(* IEC 61131-3 sources: NachHouse_TST/ROOM_API_PILOT/CODEX_BACKUP_BEFORE_SK_COMMENTS_20260826_2356, 11 files *)

(* ---- 02_TYPES.ST ---- *)
(* ROOM_API_PILOT - logical API and transport types. *)

TYPE T_API_COMMAND_RESULT :
STRUCT
    ClientId       : STRING[36];
    RequestId      : UDINT;
    Result         : USINT;
    Message        : STRING[80];
    ConfigRevision : UDINT;
    StateRevision  : UDINT;
END_STRUCT
END_TYPE

TYPE T_API_INFO :
STRUCT
    ApiVersion        : STRING[32];
    ConfigRevision    : UDINT;
    StateRevision     : UDINT;
    MaxRooms          : USINT;
    LastCommandResult : T_API_COMMAND_RESULT;
END_STRUCT
END_TYPE

TYPE T_ROOM_CONFIG :
STRUCT
    Used        : BOOL;
    RoomId      : UDINT;
    Name        : STRING[64];
    ProjectName : STRING[64];
    IconId      : UINT;
    SortDefault : UINT;
END_STRUCT
END_TYPE

TYPE T_API_CONFIG :
STRUCT
    Rooms : ARRAY[1..40] OF T_ROOM_CONFIG;
END_STRUCT
END_TYPE

TYPE T_ROOM_STATE :
STRUCT
    RoomId       : UDINT;
    Temperature  : REAL;
    Humidity     : REAL;
    Presence     : BOOL;
    DayPhase     : UINT;
    CategoryMask : DWORD;
    AlarmLevel   : USINT;
    Online       : BOOL;
END_STRUCT
END_TYPE

TYPE T_API_STATE :
STRUCT
    Rooms : ARRAY[1..40] OF T_ROOM_STATE;
END_STRUCT
END_TYPE

TYPE T_API_COMMAND_ROOM :
STRUCT
    ClientId     : STRING[36];
    RequestId    : UDINT;
    Action       : USINT;
    RoomId       : UDINT;
    SourceRoomId : UDINT;
    Name         : STRING[64];
    ProjectName  : STRING[64];
END_STRUCT
END_TYPE

TYPE T_API_CONFIG_CHANGE :
STRUCT
    Valid     : BOOL;
    Operation : USINT;
    RoomId    : UDINT;
    Room      : T_ROOM_CONFIG;
END_STRUCT
END_TYPE

TYPE T_API_STATE_CHANGE :
STRUCT
    Valid     : BOOL;
    Operation : USINT;
    RoomId    : UDINT;
    Room      : T_ROOM_STATE;
END_STRUCT
END_TYPE

TYPE T_API_CONFIG_DIFF :
STRUCT
    Valid        : BOOL;
    FromRevision : UDINT;
    ToRevision   : UDINT;
    FullRequired : BOOL;
    ChangeCount  : USINT;
    Changes      : ARRAY[1..40] OF T_API_CONFIG_CHANGE;
END_STRUCT
END_TYPE

TYPE T_API_STATE_DIFF :
STRUCT
    Valid        : BOOL;
    FromRevision : UDINT;
    ToRevision   : UDINT;
    FullRequired : BOOL;
    ChangeCount  : USINT;
    Changes      : ARRAY[1..40] OF T_API_STATE_CHANGE;
END_STRUCT
END_TYPE

(* Transport handshake used to retrieve one retained diff frame. *)
TYPE T_API_SYNC_REQUEST :
STRUCT
    ClientId           : STRING[36];
    RequestId          : UDINT;
    ConfigFromRevision : UDINT;
    StateFromRevision  : UDINT;
END_STRUCT
END_TYPE

TYPE T_API_SYNC_RESPONSE :
STRUCT
    ClientId   : STRING[36];
    RequestId  : UDINT;
    Result     : USINT;
    Message    : STRING[80];
    ConfigMode : USINT;
    StateMode  : USINT;
    ConfigDiff : T_API_CONFIG_DIFF;
    StateDiff  : T_API_STATE_DIFF;
END_STRUCT
END_TYPE

(* Manual test input. It is deliberately separate from ApiCommand.Room. *)
TYPE T_API_TEST_STATE_REQUEST :
STRUCT
    ClientId     : STRING[36];
    RequestId    : UDINT;
    RoomId       : UDINT;
    Temperature  : REAL;
    Humidity     : REAL;
    Presence     : BOOL;
    DayPhase     : UINT;
    CategoryMask : DWORD;
    AlarmLevel   : USINT;
    Online       : BOOL;
END_STRUCT
END_TYPE

(* ---- 01_CONSTANTS.ST ---- *)
(* ROOM_API_PILOT - public numeric contract and limits. *)

VAR_GLOBAL CONSTANT
    C_API_VERSION          : STRING[32] := 'ROOM_API_PILOT/1';
    C_MAX_ROOMS            : USINT := 40;
    C_DIFF_HISTORY_DEPTH   : USINT := 8;

    API_ACTION_NONE          : USINT := 0;
    API_ACTION_ADD_ROOM      : USINT := 1;
    API_ACTION_DELETE_ROOM   : USINT := 2;
    API_ACTION_COPY_ROOM     : USINT := 3;
    API_ACTION_SET_ROOM_DATA : USINT := 4;

    API_RESULT_NONE               : USINT := 0;
    API_RESULT_OK                 : USINT := 1;
    API_RESULT_ERROR              : USINT := 2;
    API_RESULT_NOT_FOUND          : USINT := 3;
    API_RESULT_NO_FREE_SLOT       : USINT := 4;
    API_RESULT_ALREADY_EXISTS     : USINT := 5;
    API_RESULT_INVALID_ARGUMENT   : USINT := 6;
    API_RESULT_UNSUPPORTED_ACTION : USINT := 7;

    API_DIFF_NONE   : USINT := 0;
    API_DIFF_UPSERT : USINT := 1;
    API_DIFF_DELETE : USINT := 2;

    API_SYNC_CURRENT       : USINT := 0;
    API_SYNC_DIFF          : USINT := 1;
    API_SYNC_FULL_REQUIRED : USINT := 2;

    API_ALARM_OK      : USINT := 0;
    API_ALARM_WARNING : USINT := 1;
    API_ALARM_ALARM   : USINT := 2;

    API_DAY_PHASE_DAY   : UINT := 140;
    API_DAY_PHASE_DUSK  : UINT := 142;
    API_DAY_PHASE_NIGHT : UINT := 144;
    API_DAY_PHASE_DAWN  : UINT := 146;

    API_DEFAULT_ICON_ID     : UINT := 16;
    API_DEFAULT_TEMPERATURE : REAL := 20.0;
    API_DEFAULT_HUMIDITY    : REAL := 40.0;
END_VAR

(* ---- 03_PUBLIC_API.ST ---- *)
(*
   All client-visible objects are global and marked PUBLIC_API.
   The client must write request payload fields first and Execute last.
   Snapshot objects ApiConfig and ApiState are read-only by contract.
*)

VAR_GLOBAL
    ApiInfo       {PUBLIC_API} : T_API_INFO;
    ApiConfig     {PUBLIC_API} : T_API_CONFIG;
    ApiState      {PUBLIC_API} : T_API_STATE;

    ApiConfigDiff {PUBLIC_API} : T_API_CONFIG_DIFF;
    ApiStateDiff  {PUBLIC_API} : T_API_STATE_DIFF;

    ApiCommandRoom     {PUBLIC_API} : T_API_COMMAND_ROOM;
    ApiCommandExecute  {PUBLIC_API} : BOOL;
    ApiCommandBusy     {PUBLIC_API} : BOOL;
    ApiCommandFinished {PUBLIC_API} : BOOL;
    ApiCommandResult   {PUBLIC_API} : T_API_COMMAND_RESULT;

    ApiSyncRequest  {PUBLIC_API} : T_API_SYNC_REQUEST;
    ApiSyncExecute  {PUBLIC_API} : BOOL;
    ApiSyncBusy     {PUBLIC_API} : BOOL;
    ApiSyncFinished {PUBLIC_API} : BOOL;
    ApiSyncResponse {PUBLIC_API} : T_API_SYNC_RESPONSE;

    ApiTestStateRequest  {PUBLIC_API} : T_API_TEST_STATE_REQUEST;
    ApiTestStateExecute  {PUBLIC_API} : BOOL;
    ApiTestStateBusy     {PUBLIC_API} : BOOL;
    ApiTestStateFinished {PUBLIC_API} : BOOL;
    ApiTestStateResult   {PUBLIC_API} : T_API_COMMAND_RESULT;
END_VAR

(* ---- 04_INTERNAL.ST ---- *)
(* Internal state is not exported to TecoApi / PLCComS. *)

VAR_GLOBAL
    ApiInitialized : BOOL;

    ApiConfigShadow : ARRAY[1..40] OF T_ROOM_CONFIG;
    ApiStateShadow  : ARRAY[1..40] OF T_ROOM_STATE;

    ApiConfigDiffHistory : ARRAY[1..8] OF T_API_CONFIG_DIFF;
    ApiStateDiffHistory  : ARRAY[1..8] OF T_API_STATE_DIFF;
    ApiConfigHistoryHead : USINT;
    ApiStateHistoryHead  : USINT;

    ApiLastCommandClientId  : STRING[36];
    ApiLastCommandRequestId : UDINT;
    ApiLastStoredResult     : T_API_COMMAND_RESULT;
END_VAR

(* ---- 05_UTILS.ST ---- *)
(* ROOM_API_PILOT - small deterministic helpers. *)

FUNCTION ApiRoomConfigEqual : BOOL
VAR_INPUT
    A : T_ROOM_CONFIG;
    B : T_ROOM_CONFIG;
END_VAR

ApiRoomConfigEqual :=
    (A.Used = B.Used) AND
    (A.RoomId = B.RoomId) AND
    (A.Name = B.Name) AND
    (A.ProjectName = B.ProjectName) AND
    (A.IconId = B.IconId) AND
    (A.SortDefault = B.SortDefault);
END_FUNCTION

FUNCTION ApiRoomStateEqual : BOOL
VAR_INPUT
    A : T_ROOM_STATE;
    B : T_ROOM_STATE;
END_VAR

ApiRoomStateEqual :=
    (A.RoomId = B.RoomId) AND
    (A.Temperature = B.Temperature) AND
    (A.Humidity = B.Humidity) AND
    (A.Presence = B.Presence) AND
    (A.DayPhase = B.DayPhase) AND
    (A.CategoryMask = B.CategoryMask) AND
    (A.AlarmLevel = B.AlarmLevel) AND
    (A.Online = B.Online);
END_FUNCTION

FUNCTION ApiFindConfigSlot : USINT
VAR_INPUT
    RoomId : UDINT;
END_VAR
VAR
    i : USINT;
END_VAR

ApiFindConfigSlot := 0;
IF RoomId <> 0 THEN
    FOR i := 1 TO C_MAX_ROOMS DO
        IF ApiConfig.Rooms[i].Used AND (ApiConfig.Rooms[i].RoomId = RoomId) THEN
            ApiFindConfigSlot := i;
            RETURN;
        END_IF;
    END_FOR;
END_IF;
END_FUNCTION

FUNCTION ApiFindStateSlot : USINT
VAR_INPUT
    RoomId : UDINT;
END_VAR
VAR
    i : USINT;
END_VAR

ApiFindStateSlot := 0;
IF RoomId <> 0 THEN
    FOR i := 1 TO C_MAX_ROOMS DO
        IF ApiState.Rooms[i].RoomId = RoomId THEN
            ApiFindStateSlot := i;
            RETURN;
        END_IF;
    END_FOR;
END_IF;
END_FUNCTION

FUNCTION ApiFindFreeConfigSlot : USINT
VAR
    i : USINT;
END_VAR

ApiFindFreeConfigSlot := 0;
FOR i := 1 TO C_MAX_ROOMS DO
    IF NOT ApiConfig.Rooms[i].Used THEN
        ApiFindFreeConfigSlot := i;
        RETURN;
    END_IF;
END_FOR;
END_FUNCTION

FUNCTION ApiFindFreeStateSlot : USINT
VAR
    i : USINT;
END_VAR

ApiFindFreeStateSlot := 0;
FOR i := 1 TO C_MAX_ROOMS DO
    IF ApiState.Rooms[i].RoomId = 0 THEN
        ApiFindFreeStateSlot := i;
        RETURN;
    END_IF;
END_FOR;
END_FUNCTION

FUNCTION ApiClearRoomConfig : BOOL
VAR_IN_OUT
    Room : T_ROOM_CONFIG;
END_VAR

Room.Used := FALSE;
Room.RoomId := 0;
Room.Name := '';
Room.ProjectName := '';
Room.IconId := 0;
Room.SortDefault := 0;
ApiClearRoomConfig := TRUE;
END_FUNCTION

FUNCTION ApiClearRoomState : BOOL
VAR_IN_OUT
    Room : T_ROOM_STATE;
END_VAR

Room.RoomId := 0;
Room.Temperature := 0.0;
Room.Humidity := 0.0;
Room.Presence := FALSE;
Room.DayPhase := API_DAY_PHASE_DAY;
Room.CategoryMask := DWORD#16#00000000;
Room.AlarmLevel := API_ALARM_OK;
Room.Online := FALSE;
ApiClearRoomState := TRUE;
END_FUNCTION

FUNCTION ApiClearConfigDiff : BOOL
VAR_IN_OUT
    Diff : T_API_CONFIG_DIFF;
END_VAR
VAR
    i : USINT;
END_VAR

Diff.Valid := FALSE;
Diff.FromRevision := 0;
Diff.ToRevision := 0;
Diff.FullRequired := FALSE;
Diff.ChangeCount := 0;
FOR i := 1 TO C_MAX_ROOMS DO
    Diff.Changes[i].Valid := FALSE;
    Diff.Changes[i].Operation := API_DIFF_NONE;
    Diff.Changes[i].RoomId := 0;
    ApiClearRoomConfig(Diff.Changes[i].Room);
END_FOR;
ApiClearConfigDiff := TRUE;
END_FUNCTION

FUNCTION ApiClearStateDiff : BOOL
VAR_IN_OUT
    Diff : T_API_STATE_DIFF;
END_VAR
VAR
    i : USINT;
END_VAR

Diff.Valid := FALSE;
Diff.FromRevision := 0;
Diff.ToRevision := 0;
Diff.FullRequired := FALSE;
Diff.ChangeCount := 0;
FOR i := 1 TO C_MAX_ROOMS DO
    Diff.Changes[i].Valid := FALSE;
    Diff.Changes[i].Operation := API_DIFF_NONE;
    Diff.Changes[i].RoomId := 0;
    ApiClearRoomState(Diff.Changes[i].Room);
END_FOR;
ApiClearStateDiff := TRUE;
END_FUNCTION

FUNCTION ApiNextRevision : UDINT
VAR_INPUT
    Revision : UDINT;
END_VAR

ApiNextRevision := Revision + 1;
IF ApiNextRevision = 0 THEN
    ApiNextRevision := 1;
END_IF;
END_FUNCTION

FUNCTION ApiValidDayPhase : BOOL
VAR_INPUT
    DayPhase : UINT;
END_VAR

ApiValidDayPhase :=
    (DayPhase = API_DAY_PHASE_DAY) OR
    (DayPhase = API_DAY_PHASE_DUSK) OR
    (DayPhase = API_DAY_PHASE_NIGHT) OR
    (DayPhase = API_DAY_PHASE_DAWN);
END_FUNCTION

(* ---- 06_DIFF_ENGINE.ST ---- *)
(*
   Diff engine.
   One PLC transaction creates one revision and one complete diff frame.
   Eight frames are retained. A client asks for one next frame at a time.
*)

FUNCTION ApiCaptureConfigChanges : BOOL
VAR
    i          : USINT;
    count      : USINT;
    oldRev     : UDINT;
    newRev     : UDINT;
    anyChanged : BOOL;
END_VAR

anyChanged := FALSE;
FOR i := 1 TO C_MAX_ROOMS DO
    IF NOT ApiRoomConfigEqual(ApiConfig.Rooms[i], ApiConfigShadow[i]) THEN
        anyChanged := TRUE;
    END_IF;
END_FOR;

ApiCaptureConfigChanges := anyChanged;
IF NOT anyChanged THEN
    RETURN;
END_IF;

ApiClearConfigDiff(ApiConfigDiff);
oldRev := ApiInfo.ConfigRevision;
newRev := ApiNextRevision(oldRev);
ApiConfigDiff.FromRevision := oldRev;
ApiConfigDiff.ToRevision := newRev;
ApiConfigDiff.FullRequired := FALSE;
count := 0;

FOR i := 1 TO C_MAX_ROOMS DO
    IF NOT ApiRoomConfigEqual(ApiConfig.Rooms[i], ApiConfigShadow[i]) THEN
        count := count + 1;
        ApiConfigDiff.Changes[count].Valid := TRUE;

        IF ApiConfig.Rooms[i].Used THEN
            ApiConfigDiff.Changes[count].Operation := API_DIFF_UPSERT;
            ApiConfigDiff.Changes[count].RoomId := ApiConfig.Rooms[i].RoomId;
            ApiConfigDiff.Changes[count].Room := ApiConfig.Rooms[i];
        ELSE
            ApiConfigDiff.Changes[count].Operation := API_DIFF_DELETE;
            ApiConfigDiff.Changes[count].RoomId := ApiConfigShadow[i].RoomId;
            ApiClearRoomConfig(ApiConfigDiff.Changes[count].Room);
        END_IF;
    END_IF;

    ApiConfigShadow[i] := ApiConfig.Rooms[i];
END_FOR;

ApiConfigDiff.ChangeCount := count;
ApiConfigDiff.Valid := TRUE;
ApiInfo.ConfigRevision := newRev;

IF ApiConfigHistoryHead >= C_DIFF_HISTORY_DEPTH THEN
    ApiConfigHistoryHead := 1;
ELSE
    ApiConfigHistoryHead := ApiConfigHistoryHead + 1;
END_IF;
ApiConfigDiffHistory[ApiConfigHistoryHead] := ApiConfigDiff;
END_FUNCTION

FUNCTION ApiCaptureStateChanges : BOOL
VAR
    i          : USINT;
    count      : USINT;
    oldRev     : UDINT;
    newRev     : UDINT;
    anyChanged : BOOL;
END_VAR

anyChanged := FALSE;
FOR i := 1 TO C_MAX_ROOMS DO
    IF NOT ApiRoomStateEqual(ApiState.Rooms[i], ApiStateShadow[i]) THEN
        anyChanged := TRUE;
    END_IF;
END_FOR;

ApiCaptureStateChanges := anyChanged;
IF NOT anyChanged THEN
    RETURN;
END_IF;

ApiClearStateDiff(ApiStateDiff);
oldRev := ApiInfo.StateRevision;
newRev := ApiNextRevision(oldRev);
ApiStateDiff.FromRevision := oldRev;
ApiStateDiff.ToRevision := newRev;
ApiStateDiff.FullRequired := FALSE;
count := 0;

FOR i := 1 TO C_MAX_ROOMS DO
    IF NOT ApiRoomStateEqual(ApiState.Rooms[i], ApiStateShadow[i]) THEN
        count := count + 1;
        ApiStateDiff.Changes[count].Valid := TRUE;

        IF ApiState.Rooms[i].RoomId <> 0 THEN
            ApiStateDiff.Changes[count].Operation := API_DIFF_UPSERT;
            ApiStateDiff.Changes[count].RoomId := ApiState.Rooms[i].RoomId;
            ApiStateDiff.Changes[count].Room := ApiState.Rooms[i];
        ELSE
            ApiStateDiff.Changes[count].Operation := API_DIFF_DELETE;
            ApiStateDiff.Changes[count].RoomId := ApiStateShadow[i].RoomId;
            ApiClearRoomState(ApiStateDiff.Changes[count].Room);
        END_IF;
    END_IF;

    ApiStateShadow[i] := ApiState.Rooms[i];
END_FOR;

ApiStateDiff.ChangeCount := count;
ApiStateDiff.Valid := TRUE;
ApiInfo.StateRevision := newRev;

IF ApiStateHistoryHead >= C_DIFF_HISTORY_DEPTH THEN
    ApiStateHistoryHead := 1;
ELSE
    ApiStateHistoryHead := ApiStateHistoryHead + 1;
END_IF;
ApiStateDiffHistory[ApiStateHistoryHead] := ApiStateDiff;
END_FUNCTION

(* ---- 07_INIT.ST ---- *)
(* Cold-start initialization and deterministic pilot data. *)

FUNCTION ApiPilotInit : BOOL
VAR
    i : USINT;
END_VAR

ApiPilotInit := ApiInitialized;
IF ApiInitialized THEN
    RETURN;
END_IF;

FOR i := 1 TO C_MAX_ROOMS DO
    ApiClearRoomConfig(ApiConfig.Rooms[i]);
    ApiClearRoomState(ApiState.Rooms[i]);
    ApiClearRoomConfig(ApiConfigShadow[i]);
    ApiClearRoomState(ApiStateShadow[i]);
END_FOR;

FOR i := 1 TO C_DIFF_HISTORY_DEPTH DO
    ApiClearConfigDiff(ApiConfigDiffHistory[i]);
    ApiClearStateDiff(ApiStateDiffHistory[i]);
END_FOR;

(* Four sample rooms. Values are test data only. *)
ApiConfig.Rooms[1].Used := TRUE;
ApiConfig.Rooms[1].RoomId := 1;
ApiConfig.Rooms[1].Name := 'Obyvacka';
ApiConfig.Rooms[1].ProjectName := '1.01';
ApiConfig.Rooms[1].IconId := 16;
ApiConfig.Rooms[1].SortDefault := 1;

ApiConfig.Rooms[2].Used := TRUE;
ApiConfig.Rooms[2].RoomId := 2;
ApiConfig.Rooms[2].Name := 'Kuchyna';
ApiConfig.Rooms[2].ProjectName := '1.07';
ApiConfig.Rooms[2].IconId := 16;
ApiConfig.Rooms[2].SortDefault := 2;

ApiConfig.Rooms[3].Used := TRUE;
ApiConfig.Rooms[3].RoomId := 3;
ApiConfig.Rooms[3].Name := 'Spalna';
ApiConfig.Rooms[3].ProjectName := '1.09';
ApiConfig.Rooms[3].IconId := 16;
ApiConfig.Rooms[3].SortDefault := 3;

ApiConfig.Rooms[4].Used := TRUE;
ApiConfig.Rooms[4].RoomId := 4;
ApiConfig.Rooms[4].Name := 'Terasa';
ApiConfig.Rooms[4].ProjectName := 'E.01';
ApiConfig.Rooms[4].IconId := 19;
ApiConfig.Rooms[4].SortDefault := 4;

ApiState.Rooms[1].RoomId := 1;
ApiState.Rooms[1].Temperature := 22.5;
ApiState.Rooms[1].Humidity := 45.0;
ApiState.Rooms[1].Presence := TRUE;
ApiState.Rooms[1].DayPhase := API_DAY_PHASE_DAY;
ApiState.Rooms[1].CategoryMask := DWORD#16#00000007;
ApiState.Rooms[1].AlarmLevel := API_ALARM_OK;
ApiState.Rooms[1].Online := TRUE;

ApiState.Rooms[2].RoomId := 2;
ApiState.Rooms[2].Temperature := 23.0;
ApiState.Rooms[2].Humidity := 48.0;
ApiState.Rooms[2].Presence := FALSE;
ApiState.Rooms[2].DayPhase := API_DAY_PHASE_DUSK;
ApiState.Rooms[2].CategoryMask := DWORD#16#00000003;
ApiState.Rooms[2].AlarmLevel := API_ALARM_WARNING;
ApiState.Rooms[2].Online := TRUE;

ApiState.Rooms[3].RoomId := 3;
ApiState.Rooms[3].Temperature := 21.8;
ApiState.Rooms[3].Humidity := 42.0;
ApiState.Rooms[3].Presence := TRUE;
ApiState.Rooms[3].DayPhase := API_DAY_PHASE_NIGHT;
ApiState.Rooms[3].CategoryMask := DWORD#16#00000001;
ApiState.Rooms[3].AlarmLevel := API_ALARM_OK;
ApiState.Rooms[3].Online := TRUE;

ApiState.Rooms[4].RoomId := 4;
ApiState.Rooms[4].Temperature := 18.4;
ApiState.Rooms[4].Humidity := 58.0;
ApiState.Rooms[4].Presence := FALSE;
ApiState.Rooms[4].DayPhase := API_DAY_PHASE_DAWN;
ApiState.Rooms[4].CategoryMask := DWORD#16#00000004;
ApiState.Rooms[4].AlarmLevel := API_ALARM_ALARM;
ApiState.Rooms[4].Online := FALSE;

FOR i := 1 TO C_MAX_ROOMS DO
    ApiConfigShadow[i] := ApiConfig.Rooms[i];
    ApiStateShadow[i] := ApiState.Rooms[i];
END_FOR;

ApiInfo.ApiVersion := C_API_VERSION;
ApiInfo.ConfigRevision := 1;
ApiInfo.StateRevision := 1;
ApiInfo.MaxRooms := C_MAX_ROOMS;
ApiInfo.LastCommandResult.ClientId := '';
ApiInfo.LastCommandResult.RequestId := 0;
ApiInfo.LastCommandResult.Result := API_RESULT_NONE;
ApiInfo.LastCommandResult.Message := 'Ziadny prikaz';
ApiInfo.LastCommandResult.ConfigRevision := 1;
ApiInfo.LastCommandResult.StateRevision := 1;

ApiClearConfigDiff(ApiConfigDiff);
ApiConfigDiff.Valid := TRUE;
ApiConfigDiff.FromRevision := 0;
ApiConfigDiff.ToRevision := 1;
ApiConfigDiff.FullRequired := TRUE;

ApiClearStateDiff(ApiStateDiff);
ApiStateDiff.Valid := TRUE;
ApiStateDiff.FromRevision := 0;
ApiStateDiff.ToRevision := 1;
ApiStateDiff.FullRequired := TRUE;

ApiCommandRoom.ClientId := '';
ApiCommandRoom.RequestId := 0;
ApiCommandRoom.Action := API_ACTION_NONE;
ApiCommandRoom.RoomId := 0;
ApiCommandRoom.SourceRoomId := 0;
ApiCommandRoom.Name := '';
ApiCommandRoom.ProjectName := '';
ApiCommandExecute := FALSE;
ApiCommandBusy := FALSE;
ApiCommandFinished := FALSE;
ApiCommandResult := ApiInfo.LastCommandResult;

ApiSyncExecute := FALSE;
ApiSyncBusy := FALSE;
ApiSyncFinished := FALSE;
ApiTestStateExecute := FALSE;
ApiTestStateBusy := FALSE;
ApiTestStateFinished := FALSE;

ApiConfigHistoryHead := 0;
ApiStateHistoryHead := 0;
ApiLastCommandClientId := '';
ApiLastCommandRequestId := 0;
ApiLastStoredResult := ApiInfo.LastCommandResult;

ApiInitialized := TRUE;
ApiPilotInit := TRUE;
END_FUNCTION

(* ---- 08_COMMAND_ENGINE.ST ---- *)
(* ADD / DELETE / COPY / SET command processor. *)

FUNCTION ApiProcessRoomCommand : BOOL
VAR
    i             : USINT;
    configSlot    : USINT;
    stateSlot     : USINT;
    sourceCfgSlot : USINT;
    sourceStSlot  : USINT;
    maxSort       : UINT;
    sourceSort    : UINT;
    resultCode    : USINT;
    resultMessage : STRING[80];
    executeChange : BOOL;
END_VAR

ApiProcessRoomCommand := FALSE;
IF NOT ApiCommandExecute THEN
    RETURN;
END_IF;

ApiProcessRoomCommand := TRUE;
ApiCommandBusy := TRUE;
ApiCommandFinished := FALSE;

(* Exact retry of the latest command is idempotent. *)
IF (ApiCommandRoom.ClientId = ApiLastCommandClientId) AND
   (ApiCommandRoom.RequestId = ApiLastCommandRequestId) AND
   (ApiCommandRoom.RequestId <> 0) THEN

    ApiCommandResult := ApiLastStoredResult;
    ApiInfo.LastCommandResult := ApiLastStoredResult;

ELSE
    resultCode := API_RESULT_OK;
    resultMessage := 'OK';
    executeChange := FALSE;

    IF (ApiCommandRoom.ClientId = '') OR (ApiCommandRoom.RequestId = 0) THEN
        resultCode := API_RESULT_INVALID_ARGUMENT;
        resultMessage := 'Neplatny ClientId alebo RequestId';
    ELSE
        CASE ApiCommandRoom.Action OF

            API_ACTION_ADD_ROOM:
                IF (ApiCommandRoom.RoomId = 0) OR (ApiCommandRoom.Name = '') THEN
                    resultCode := API_RESULT_INVALID_ARGUMENT;
                    resultMessage := 'Neplatne ID alebo nazov';
                ELSIF ApiFindConfigSlot(ApiCommandRoom.RoomId) <> 0 THEN
                    resultCode := API_RESULT_ALREADY_EXISTS;
                    resultMessage := 'RoomId uz existuje';
                ELSE
                    configSlot := ApiFindFreeConfigSlot();
                    stateSlot := ApiFindFreeStateSlot();
                    IF (configSlot = 0) OR (stateSlot = 0) THEN
                        resultCode := API_RESULT_NO_FREE_SLOT;
                        resultMessage := 'Nie je volny slot';
                    ELSE
                        maxSort := 0;
                        FOR i := 1 TO C_MAX_ROOMS DO
                            IF ApiConfig.Rooms[i].Used AND
                               (ApiConfig.Rooms[i].SortDefault > maxSort) THEN
                                maxSort := ApiConfig.Rooms[i].SortDefault;
                            END_IF;
                        END_FOR;

                        ApiClearRoomConfig(ApiConfig.Rooms[configSlot]);
                        ApiConfig.Rooms[configSlot].Used := TRUE;
                        ApiConfig.Rooms[configSlot].RoomId := ApiCommandRoom.RoomId;
                        ApiConfig.Rooms[configSlot].Name := ApiCommandRoom.Name;
                        ApiConfig.Rooms[configSlot].ProjectName := ApiCommandRoom.ProjectName;
                        ApiConfig.Rooms[configSlot].IconId := API_DEFAULT_ICON_ID;
                        ApiConfig.Rooms[configSlot].SortDefault := maxSort + 1;

                        ApiClearRoomState(ApiState.Rooms[stateSlot]);
                        ApiState.Rooms[stateSlot].RoomId := ApiCommandRoom.RoomId;
                        ApiState.Rooms[stateSlot].Temperature := API_DEFAULT_TEMPERATURE;
                        ApiState.Rooms[stateSlot].Humidity := API_DEFAULT_HUMIDITY;
                        ApiState.Rooms[stateSlot].Presence := FALSE;
                        ApiState.Rooms[stateSlot].DayPhase := API_DAY_PHASE_DAY;
                        ApiState.Rooms[stateSlot].CategoryMask := DWORD#16#00000000;
                        ApiState.Rooms[stateSlot].AlarmLevel := API_ALARM_OK;
                        ApiState.Rooms[stateSlot].Online := TRUE;

                        executeChange := TRUE;
                        resultMessage := 'Miestnost pridana';
                    END_IF;
                END_IF;

            API_ACTION_DELETE_ROOM:
                configSlot := ApiFindConfigSlot(ApiCommandRoom.RoomId);
                stateSlot := ApiFindStateSlot(ApiCommandRoom.RoomId);
                IF (configSlot = 0) OR (stateSlot = 0) THEN
                    resultCode := API_RESULT_NOT_FOUND;
                    resultMessage := 'Miestnost nenajdena';
                ELSE
                    ApiClearRoomConfig(ApiConfig.Rooms[configSlot]);
                    ApiClearRoomState(ApiState.Rooms[stateSlot]);
                    executeChange := TRUE;
                    resultMessage := 'Miestnost zmazana';
                END_IF;

            API_ACTION_COPY_ROOM:
                sourceCfgSlot := ApiFindConfigSlot(ApiCommandRoom.SourceRoomId);
                sourceStSlot := ApiFindStateSlot(ApiCommandRoom.SourceRoomId);
                IF (ApiCommandRoom.RoomId = 0) OR
                   (ApiCommandRoom.RoomId = ApiCommandRoom.SourceRoomId) THEN
                    resultCode := API_RESULT_INVALID_ARGUMENT;
                    resultMessage := 'Neplatne cielove RoomId';
                ELSIF (sourceCfgSlot = 0) OR (sourceStSlot = 0) THEN
                    resultCode := API_RESULT_NOT_FOUND;
                    resultMessage := 'Zdrojova miestnost nenajdena';
                ELSIF ApiFindConfigSlot(ApiCommandRoom.RoomId) <> 0 THEN
                    resultCode := API_RESULT_ALREADY_EXISTS;
                    resultMessage := 'Cielove RoomId uz existuje';
                ELSE
                    configSlot := ApiFindFreeConfigSlot();
                    stateSlot := ApiFindFreeStateSlot();
                    IF (configSlot = 0) OR (stateSlot = 0) THEN
                        resultCode := API_RESULT_NO_FREE_SLOT;
                        resultMessage := 'Nie je volny slot';
                    ELSE
                        sourceSort := ApiConfig.Rooms[sourceCfgSlot].SortDefault;
                        FOR i := 1 TO C_MAX_ROOMS DO
                            IF ApiConfig.Rooms[i].Used AND
                               (ApiConfig.Rooms[i].SortDefault > sourceSort) THEN
                                ApiConfig.Rooms[i].SortDefault :=
                                    ApiConfig.Rooms[i].SortDefault + 1;
                            END_IF;
                        END_FOR;

                        ApiConfig.Rooms[configSlot] := ApiConfig.Rooms[sourceCfgSlot];
                        ApiConfig.Rooms[configSlot].RoomId := ApiCommandRoom.RoomId;
                        ApiConfig.Rooms[configSlot].SortDefault := sourceSort + 1;
                        IF ApiCommandRoom.Name <> '' THEN
                            ApiConfig.Rooms[configSlot].Name := ApiCommandRoom.Name;
                        END_IF;
                        IF ApiCommandRoom.ProjectName <> '' THEN
                            ApiConfig.Rooms[configSlot].ProjectName := ApiCommandRoom.ProjectName;
                        END_IF;

                        ApiState.Rooms[stateSlot] := ApiState.Rooms[sourceStSlot];
                        ApiState.Rooms[stateSlot].RoomId := ApiCommandRoom.RoomId;

                        executeChange := TRUE;
                        resultMessage := 'Miestnost skopirovana';
                    END_IF;
                END_IF;

            API_ACTION_SET_ROOM_DATA:
                configSlot := ApiFindConfigSlot(ApiCommandRoom.RoomId);
                IF configSlot = 0 THEN
                    resultCode := API_RESULT_NOT_FOUND;
                    resultMessage := 'Miestnost nenajdena';
                ELSIF ApiCommandRoom.Name = '' THEN
                    resultCode := API_RESULT_INVALID_ARGUMENT;
                    resultMessage := 'Nazov nesmie byt prazdny';
                ELSE
                    ApiConfig.Rooms[configSlot].Name := ApiCommandRoom.Name;
                    ApiConfig.Rooms[configSlot].ProjectName := ApiCommandRoom.ProjectName;
                    executeChange := TRUE;
                    resultMessage := 'Udaje miestnosti nastavene';
                END_IF;

            ELSE
                resultCode := API_RESULT_UNSUPPORTED_ACTION;
                resultMessage := 'Nepodporovana akcia';
        END_CASE;
    END_IF;

    IF executeChange AND (resultCode = API_RESULT_OK) THEN
        ApiCaptureConfigChanges();
        ApiCaptureStateChanges();
    END_IF;

    ApiCommandResult.ClientId := ApiCommandRoom.ClientId;
    ApiCommandResult.RequestId := ApiCommandRoom.RequestId;
    ApiCommandResult.Result := resultCode;
    ApiCommandResult.Message := resultMessage;
    ApiCommandResult.ConfigRevision := ApiInfo.ConfigRevision;
    ApiCommandResult.StateRevision := ApiInfo.StateRevision;

    ApiInfo.LastCommandResult := ApiCommandResult;
    ApiLastCommandClientId := ApiCommandRoom.ClientId;
    ApiLastCommandRequestId := ApiCommandRoom.RequestId;
    ApiLastStoredResult := ApiCommandResult;
END_IF;

ApiCommandExecute := FALSE;
ApiCommandBusy := FALSE;
ApiCommandFinished := TRUE;
END_FUNCTION

(* ---- 09_STATE_TEST.ST ---- *)
(* Manual, validated test-state writer. No real IO is connected. *)

FUNCTION ApiProcessTestState : BOOL
VAR
    configSlot    : USINT;
    stateSlot     : USINT;
    resultCode    : USINT;
    resultMessage : STRING[80];
END_VAR

ApiProcessTestState := FALSE;
IF NOT ApiTestStateExecute THEN
    RETURN;
END_IF;

ApiProcessTestState := TRUE;
ApiTestStateBusy := TRUE;
ApiTestStateFinished := FALSE;
resultCode := API_RESULT_OK;
resultMessage := 'Testovaci stav nastaveny';

configSlot := ApiFindConfigSlot(ApiTestStateRequest.RoomId);
stateSlot := ApiFindStateSlot(ApiTestStateRequest.RoomId);

IF (ApiTestStateRequest.ClientId = '') OR
   (ApiTestStateRequest.RequestId = 0) THEN
    resultCode := API_RESULT_INVALID_ARGUMENT;
    resultMessage := 'Neplatny ClientId alebo RequestId';
ELSIF (configSlot = 0) OR (stateSlot = 0) THEN
    resultCode := API_RESULT_NOT_FOUND;
    resultMessage := 'Miestnost nenajdena';
ELSIF (ApiTestStateRequest.Temperature < -50.0) OR
      (ApiTestStateRequest.Temperature > 100.0) OR
      (ApiTestStateRequest.Humidity < 0.0) OR
      (ApiTestStateRequest.Humidity > 100.0) OR
      (ApiTestStateRequest.AlarmLevel > API_ALARM_ALARM) OR
      (NOT ApiValidDayPhase(ApiTestStateRequest.DayPhase)) THEN
    resultCode := API_RESULT_INVALID_ARGUMENT;
    resultMessage := 'Neplatna testovacia hodnota';
ELSE
    ApiState.Rooms[stateSlot].Temperature := ApiTestStateRequest.Temperature;
    ApiState.Rooms[stateSlot].Humidity := ApiTestStateRequest.Humidity;
    ApiState.Rooms[stateSlot].Presence := ApiTestStateRequest.Presence;
    ApiState.Rooms[stateSlot].DayPhase := ApiTestStateRequest.DayPhase;
    ApiState.Rooms[stateSlot].CategoryMask := ApiTestStateRequest.CategoryMask;
    ApiState.Rooms[stateSlot].AlarmLevel := ApiTestStateRequest.AlarmLevel;
    ApiState.Rooms[stateSlot].Online := ApiTestStateRequest.Online;
    ApiCaptureStateChanges();
END_IF;

ApiTestStateResult.ClientId := ApiTestStateRequest.ClientId;
ApiTestStateResult.RequestId := ApiTestStateRequest.RequestId;
ApiTestStateResult.Result := resultCode;
ApiTestStateResult.Message := resultMessage;
ApiTestStateResult.ConfigRevision := ApiInfo.ConfigRevision;
ApiTestStateResult.StateRevision := ApiInfo.StateRevision;

ApiTestStateExecute := FALSE;
ApiTestStateBusy := FALSE;
ApiTestStateFinished := TRUE;
END_FUNCTION

(* ---- 10_SYNC_ENGINE.ST ---- *)
(* Cache recovery: return one next retained frame or request a full snapshot. *)

FUNCTION ApiProcessSyncRequest : BOOL
VAR
    i           : USINT;
    foundConfig : BOOL;
    foundState  : BOOL;
END_VAR

ApiProcessSyncRequest := FALSE;
IF NOT ApiSyncExecute THEN
    RETURN;
END_IF;

ApiProcessSyncRequest := TRUE;
ApiSyncBusy := TRUE;
ApiSyncFinished := FALSE;

ApiSyncResponse.ClientId := ApiSyncRequest.ClientId;
ApiSyncResponse.RequestId := ApiSyncRequest.RequestId;
ApiSyncResponse.Result := API_RESULT_OK;
ApiSyncResponse.Message := 'Synchronizacia pripravena';

ApiClearConfigDiff(ApiSyncResponse.ConfigDiff);
ApiClearStateDiff(ApiSyncResponse.StateDiff);
foundConfig := FALSE;
foundState := FALSE;

IF (ApiSyncRequest.ClientId = '') OR (ApiSyncRequest.RequestId = 0) THEN
    ApiSyncResponse.Result := API_RESULT_INVALID_ARGUMENT;
    ApiSyncResponse.Message := 'Neplatny ClientId alebo RequestId';
END_IF;

IF ApiSyncRequest.ConfigFromRevision = ApiInfo.ConfigRevision THEN
    ApiSyncResponse.ConfigMode := API_SYNC_CURRENT;
    ApiSyncResponse.ConfigDiff.Valid := TRUE;
    ApiSyncResponse.ConfigDiff.FromRevision := ApiInfo.ConfigRevision;
    ApiSyncResponse.ConfigDiff.ToRevision := ApiInfo.ConfigRevision;
    foundConfig := TRUE;
ELSE
    FOR i := 1 TO C_DIFF_HISTORY_DEPTH DO
        IF ApiConfigDiffHistory[i].Valid AND
           (ApiConfigDiffHistory[i].FromRevision =
            ApiSyncRequest.ConfigFromRevision) THEN
            ApiSyncResponse.ConfigDiff := ApiConfigDiffHistory[i];
            ApiSyncResponse.ConfigMode := API_SYNC_DIFF;
            foundConfig := TRUE;
            EXIT;
        END_IF;
    END_FOR;
END_IF;

IF NOT foundConfig THEN
    ApiSyncResponse.ConfigMode := API_SYNC_FULL_REQUIRED;
    ApiSyncResponse.ConfigDiff.Valid := TRUE;
    ApiSyncResponse.ConfigDiff.FromRevision := ApiSyncRequest.ConfigFromRevision;
    ApiSyncResponse.ConfigDiff.ToRevision := ApiInfo.ConfigRevision;
    ApiSyncResponse.ConfigDiff.FullRequired := TRUE;
END_IF;

IF ApiSyncRequest.StateFromRevision = ApiInfo.StateRevision THEN
    ApiSyncResponse.StateMode := API_SYNC_CURRENT;
    ApiSyncResponse.StateDiff.Valid := TRUE;
    ApiSyncResponse.StateDiff.FromRevision := ApiInfo.StateRevision;
    ApiSyncResponse.StateDiff.ToRevision := ApiInfo.StateRevision;
    foundState := TRUE;
ELSE
    FOR i := 1 TO C_DIFF_HISTORY_DEPTH DO
        IF ApiStateDiffHistory[i].Valid AND
           (ApiStateDiffHistory[i].FromRevision =
            ApiSyncRequest.StateFromRevision) THEN
            ApiSyncResponse.StateDiff := ApiStateDiffHistory[i];
            ApiSyncResponse.StateMode := API_SYNC_DIFF;
            foundState := TRUE;
            EXIT;
        END_IF;
    END_FOR;
END_IF;

IF NOT foundState THEN
    ApiSyncResponse.StateMode := API_SYNC_FULL_REQUIRED;
    ApiSyncResponse.StateDiff.Valid := TRUE;
    ApiSyncResponse.StateDiff.FromRevision := ApiSyncRequest.StateFromRevision;
    ApiSyncResponse.StateDiff.ToRevision := ApiInfo.StateRevision;
    ApiSyncResponse.StateDiff.FullRequired := TRUE;
END_IF;

ApiSyncExecute := FALSE;
ApiSyncBusy := FALSE;
ApiSyncFinished := TRUE;
END_FUNCTION

(* ---- prgMain.ST ---- *)
PROGRAM prgMain
VAR
END_VAR

ApiPilotInit();

IF ApiInitialized THEN
    ApiProcessRoomCommand();
    ApiProcessTestState();

    (* Also catches manual edits made from the Mosaic watch window. *)
    ApiCaptureConfigChanges();
    ApiCaptureStateChanges();

    ApiProcessSyncRequest();
END_IF;
END_PROGRAM
